(* IEC 61131-3 sources: ZPLC/tools/ai-eval/fixtures/st-repair/project/src, 1 file *)

(* ---- LatchTwoSensors.st ---- *)
PROGRAM LatchTwoSensors
VAR_INPUT
    EyeA AT %I0.0 : BOOL;
    EyeB AT %I0.1 : BOOL;
END_VAR
VAR_OUTPUT
    Run AT %Q0.0 : BOOL;
END_VAR

IF EyeA THEN
    Run := TRUE;
END_IF;
IF EyeB THEN
    Run := TRUE;
END_IF;

END_PROGRAM
